FUNCTION_BLOCK HeatCalc (* Basic Function Block Type *)
  (* Standard: 61499-2 *)
  (* Version 0.0, 6/21/2016, Andrei, nxtControl GmbH, Template *)
  PACKAGE Main;
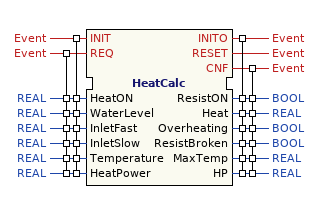
  EVENT_INPUT
    INIT WITH HeatON, WaterLevel, InletFast, InletSlow, Temperature, HeatPower; (* Initialization Request *)
    REQ WITH HeatON, WaterLevel, InletFast, InletSlow, Temperature, HeatPower; (* Normal Execution Request *)
  END_EVENT
  EVENT_OUTPUT
    INITO WITH ResistON, Heat, Overheating, ResistBroken, MaxTemp, HP; (* Initialization Confirm *)
    RESET;
    CNF WITH ResistON, Heat, Overheating, ResistBroken, MaxTemp, HP; (* Execution Confirmation *)
  END_EVENT
  VAR_INPUT
    HeatON : REAL; (* Input event qualifier *)
    WaterLevel : REAL;
    InletFast : REAL;
    InletSlow : REAL;
    Temperature : REAL;
    HeatPower : REAL;
  END_VAR
  VAR_OUTPUT
    ResistON : BOOL;
    Heat : REAL; (* Output event qualifier *)
    Overheating : BOOL;
    ResistBroken : BOOL;
    MaxTemp : REAL;
    HP : REAL;
  END_VAR
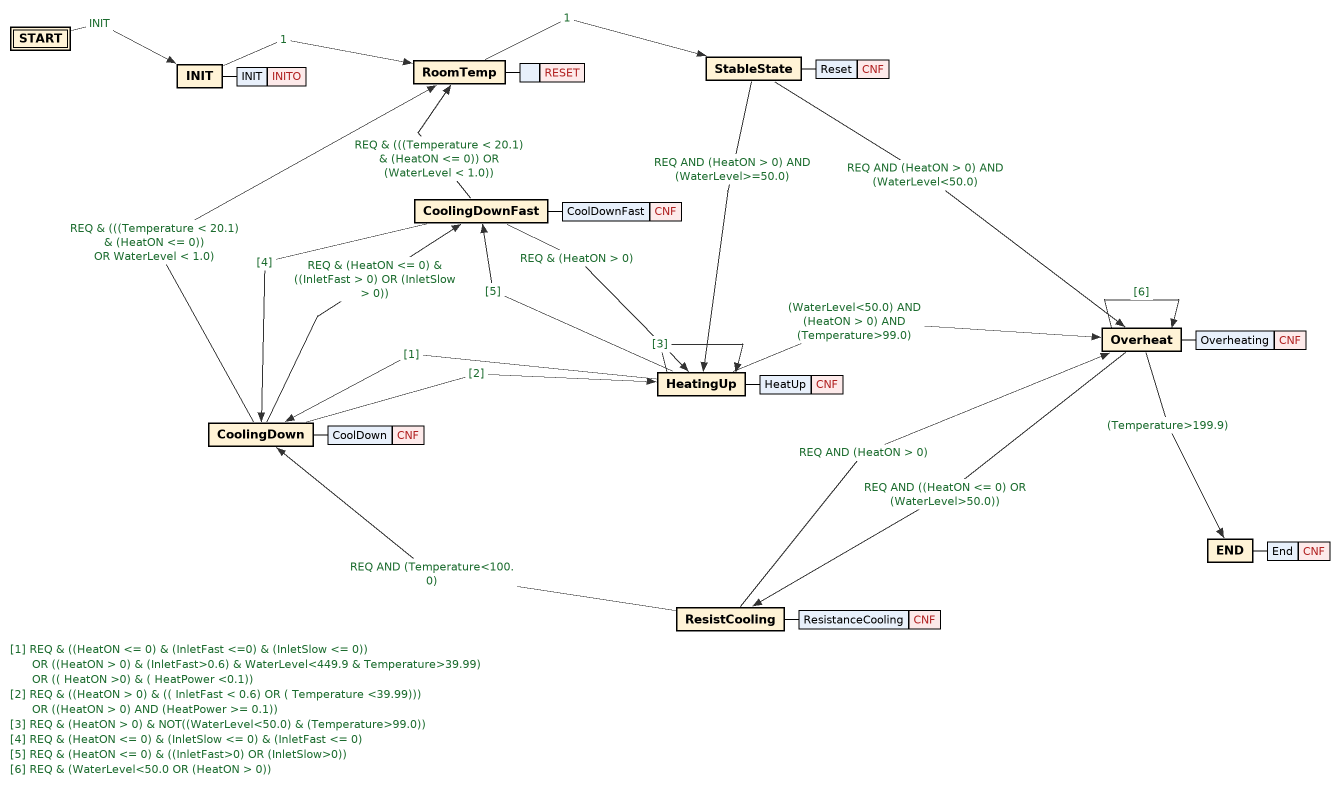
  EC_STATES
    START; (* Initial State *)
    INIT : INIT -> INITO; (* Initialization *)
    HeatingUp : HeatUp -> CNF; (* Normal execution *)
    CoolingDown : CoolDown -> CNF;
    RoomTemp : -> RESET;
    END : End -> CNF;
    StableState : Reset -> CNF;
    Overheat : Overheating -> CNF;
    ResistCooling : ResistanceCooling -> CNF;
    CoolingDownFast : CoolDownFast -> CNF;
  END_STATES
  EC_TRANSITIONS
    START TO INIT := INIT;
    INIT TO RoomTemp := 1;
    CoolingDown TO HeatingUp := REQ & ((HeatON > 0) & (( InletFast < 0.6) OR ( Temperature <39.99))) OR ((HeatON > 0) AND (HeatPower >= 0.1));
    HeatingUp TO Overheat := (WaterLevel<50.0) AND (HeatON > 0) AND (Temperature>99.0);
    RoomTemp TO StableState := 1;
    StableState TO HeatingUp := REQ AND (HeatON > 0) AND (WaterLevel>=50.0);
    CoolingDown TO RoomTemp := REQ & (((Temperature < 20.1) & (HeatON <= 0)) OR WaterLevel < 1.0);
    ResistCooling TO CoolingDown := REQ AND (Temperature<100.0);
    Overheat TO END := (Temperature>199.9);
    Overheat TO ResistCooling := REQ AND ((HeatON <= 0) OR (WaterLevel>50.0));
    ResistCooling TO Overheat := REQ AND (HeatON > 0);
    StableState TO Overheat := REQ AND (HeatON > 0) AND (WaterLevel<50.0);
    CoolingDownFast TO RoomTemp := REQ & (((Temperature < 20.1) & (HeatON <= 0)) OR (WaterLevel < 1.0));
    HeatingUp TO CoolingDownFast := REQ & (HeatON <= 0) & ((InletFast>0) OR (InletSlow>0));
    CoolingDownFast TO CoolingDown := REQ & (HeatON <= 0) & (InletSlow <= 0) & (InletFast <= 0);
    CoolingDownFast TO HeatingUp := REQ & (HeatON > 0);
    CoolingDown TO CoolingDownFast := REQ & (HeatON <= 0) & ((InletFast > 0) OR (InletSlow > 0));
    HeatingUp TO HeatingUp := REQ & (HeatON > 0) & NOT((WaterLevel<50.0) & (Temperature>99.0));
    Overheat TO Overheat := REQ & (WaterLevel<50.0 OR (HeatON > 0));
    HeatingUp TO CoolingDown := REQ & ((HeatON <= 0) & (InletFast <=0) & (InletSlow <= 0)) OR ((HeatON > 0) & (InletFast>0.6) & WaterLevel<449.9 & Temperature>39.99) OR (( HeatON >0) & ( HeatPower <0.1));
  END_TRANSITIONS
  ALGORITHM INIT IN ST: (* Initialization algorithm *)
Heat := 0.0;
ResistON := FALSE;
ResistBroken := FALSE;
MaxTemp := 100.0;
HP := HeatPower;
  END_ALGORITHM
  ALGORITHM HeatUp IN ST: (* Normally executed algorithm *)
Heat := HeatON*HeatPower*(450.0/(WaterLevel+50));
ResistON := TRUE;
HP := HeatPower;
  END_ALGORITHM
  ALGORITHM CoolDown IN ST:
Heat := -15;
MaxTemp := 100.0;
ResistON := FALSE;
ResistON := INT_TO_BOOL(REAL_TO_INT(HeatON));
HP := HeatPower;
  END_ALGORITHM
  ALGORITHM Reset IN ST:
Heat := 0.0;
ResistON := FALSE;
HP := HeatPower;
  END_ALGORITHM
  ALGORITHM End IN ST:
Overheating := FALSE;
ResistON := FALSE;
ResistBroken := TRUE;
Heat := -15.0;
HP := HeatPower;
  END_ALGORITHM
  ALGORITHM Overheating IN ST:
Heat := 100.0;
MaxTemp := 200.0;
ResistON := TRUE;
Overheating := TRUE;
HP := HeatPower;
  END_ALGORITHM
  ALGORITHM ResistanceCooling IN ST:
Heat := -30.0;
ResistON := TRUE;
Overheating := FALSE;
HP := HeatPower;
  END_ALGORITHM
  ALGORITHM CoolDownFast IN ST:
Heat := -30.0;
MaxTemp := 100.0;
ResistON := FALSE;
HP := HeatPower;
  END_ALGORITHM
END_FUNCTION_BLOCK
